(* IEC 61131-3 sources: Lasal-MCP/examples/SampleSource/LASALScreenAdvancedSolution/LASALScreenAdvancedSolution/LASALScreenAdvacnedSolution/Stations/Terminal/HMI/Network/CarouselNet, 1 file *)

(* ---- ONE_CarouselNet_Table.st ---- *)
#define OBJECTS_CONFIG

#include <.\lsl_st_mt.h>
//Define part of class MyCarousel
#define MAX_ITEMS 20

//***** Parameters for Carousel *****
#define HORIZONTAL_DRAW_ORDER_CARO FALSE
#define INFINITE_CARO FALSE
#define ELEMENT_GAP_CARO 5
#define FRAMEWORK_NEW_AGE_DARK 81 // ID in LSE
#define VERTICAL_SCROLL_BAR TRUE

FUNCTION GLOBAL TAB ONE_CarouselNet
-1$UINT, 0$UINT,
0$UINT, 0$UINT,

7$UDINT,
TO_UDINT(3599188277), "_Screen", 0$UINT, 3$UINT, 0$UINT,
TO_UDINT(2225119864), "MerkerEx", 1$UINT, 22$UINT, 0$UINT,
TO_UDINT(3908638574), "MyCarousel", 0$UINT, 0$UINT, 1$UINT,
TO_UDINT(933570811), "RAMex", 1$UINT, 17$UINT, 2$UINT,
TO_UDINT(2898603620), "StringInternal", 1$UINT, 84$UINT, 0$UINT,
TO_UDINT(2408581120), "StringRAM", 1$UINT, 10$UINT, 2$UINT,
TO_UDINT(3232495061), "VirtualBaseInit", 1$UINT, 3$UINT, 0$UINT,

_NO_ATTR, TO_UDINT(691952383), "MYCAROUSEL1",

1$UINT, TO_UDINT(1583852022), "MYCAROUSEL1\LASALOBJNAME\DATABUFFER",
1$UINT, TO_UDINT(547120993), "MYCAROUSEL1\LSEOBJNAME\DATABUFFER",

1$UINT, TO_UDINT(3532119425), "MYCAROUSEL1\LASALOBJNAME",
1$UINT, TO_UDINT(2829249980), "MYCAROUSEL1\LSEOBJNAME",

//Internal connections
0$UDINT,
4$UDINT,
TO_UDINT(0), "LasalObjName", TO_UDINT(3),
TO_UDINT(0), "LSEObjName", TO_UDINT(4),
TO_UDINT(3), "DataBuffer", TO_UDINT(1),
TO_UDINT(4), "DataBuffer", TO_UDINT(2),
0$UDINT,
2$UDINT,
TO_UDINT(3), "DataBuffer", TO_UDINT(1), "m_udLength",
TO_UDINT(4), "DataBuffer", TO_UDINT(2), "m_udLength",

//Initialization values
0$UDINT,
11$UDINT,
TO_UDINT(0), "xy1x", TO_UDINT(140),//|CarouselNet.MyCarousel1.xy1x;
TO_UDINT(0), "xy1y", TO_UDINT(90),//|CarouselNet.MyCarousel1.xy1y;
TO_UDINT(0), "xy2x", TO_UDINT(659),//|CarouselNet.MyCarousel1.xy2x;
TO_UDINT(0), "xy2y", TO_UDINT(454),//|CarouselNet.MyCarousel1.xy2y;
TO_UDINT(0), "Lse", TO_UDINT(0),//|CarouselNet.MyCarousel1.Lse;
TO_UDINT(0), "No", TO_UDINT(8),//|CarouselNet.MyCarousel1.No;
TO_UDINT(0), "ImA", TO_UDINT(0),//|CarouselNet.MyCarousel1.ImA;
TO_UDINT(1), "ThreadSafe", TO_UDINT(0),//|CarouselNet.LasalObjName\MyCarousel1\DataBuffer.ThreadSafe;
TO_UDINT(2), "ThreadSafe", TO_UDINT(0),//|CarouselNet.LSEObjName\MyCarousel1\DataBuffer.ThreadSafe;
TO_UDINT(3), "SingleRealloc", TO_UDINT(1),//|CarouselNet.MyCarousel1\LasalObjName.SingleRealloc;
TO_UDINT(4), "SingleRealloc", TO_UDINT(1),//|CarouselNet.MyCarousel1\LSEObjName.SingleRealloc;

//Symbolic initialization values
0$UDINT,
0$UDINT,

//Initialization of string values
0$UDINT,
2$UDINT,
TO_UDINT(3), "", 0$UINT, TO_UINT(OFF(L1)-OFF(L0)), L0:"MyValues",L1://|CarouselNet.MyCarousel1\LasalObjName.Data;
TO_UDINT(4), "", 0$UINT, TO_UINT(OFF(L3)-OFF(L2)), L2:"Value",L3://|CarouselNet.MyCarousel1\LSEObjName.Data;

//Configuration of tasks (RealTime, Cyclic, Background)
0$UDINT,
0$UDINT,

0$UDINT,
0$UDINT,

0$UDINT,
0$UDINT,

//External connections
0$UDINT,
1$UDINT,
TO_UDINT(0), "Lse", C_DIR, TO_UDINT(299963966), "Lse","Lse",

//Magic internal connections
0$UDINT,
2$UDINT,
TO_UDINT(1), "UseFile", TO_UDINT(3), "UseFile",
TO_UDINT(2), "UseFile", TO_UDINT(4), "UseFile",

//Configuration of timeslots of tasks (RealTime, Cyclic)
#ifdef __LSLLDR_TIMESLOTS__
0$UDINT,
0$UDINT,

0$UDINT,
0$UDINT,

#endif //__LSLLDR_TIMESLOTS__

//MultiMaster connections
#ifdef __LSLLDR_MULTIMASTER__
0$UDINT,
0$UDINT,
#endif //__LSLLDR_MULTIMASTER__

//Configuration for task ID (RealTime, CyclicTime)
#ifdef __LSLLDR_TASKID__
"\\\\TASKS2  "
0$UDINT,
0$UDINT,

0$UDINT,
0$UDINT,

0$UDINT,
0$UDINT,

#endif //__LSLLDR_TASKID__

END_FUNCTION
